Staubli VAL3: IOcomment.pgx

public program IOcomment(num x_nType, num x_nIndex, string x_sComment)
begin
  switch x_nType
    case 0
      io:dInItem[x_nIndex].sComment=x_sComment
      io:sCommentDin[x_nIndex]=x_sComment
    break
    case 1
      io:dOutItem[x_nIndex].sComment=x_sComment
      io:sCommentDout[x_nIndex]=x_sComment
    break
    case 2
      io:aInItem[x_nIndex].sComment=x_sComment
      io:sCommentAin[x_nIndex]=x_sComment
    break
    case 3
      io:aOutItem[x_nIndex].sComment=x_sComment
      io:sCommentAout[x_nIndex]=x_sComment
    break

  endSwitch

  io:libSave()
  delay(0)
end
